(*
SPDX-FileCopyrightText: © 2026 Oleksandr Tiutyk <trofimich@gmail.com>
SPDX-License-Identifier: MIT
License: https://opensource.org/license/mit
*)

(*!
<summary>Checks that a configured task name survives the STOPPED to READY reset.</summary>
<description>
Completes a resource-free one-step task before invoking Reset. A new local fixture is used on every run.
</description>
*)

{attribute 'no_explicit_call' := 'do not call this function block directly'}
FUNCTION_BLOCK TaskNamePreservedByResetTest EXTENDS TOF_Testing.SingleCycleTest
VAR_STAT
	{attribute 'hide'}
	_ClassName : STRING := __POUNAME();
END_VAR

//! <summary>Verifies the constructor name and exercises Reset from STOPPED before checking that name again.</summary>
METHOD PROTECTED ExecuteTest
VAR
	task : CounterTask(name := "Configured counter");
	started : BOOL;
	resetSucceeded : BOOL;
END_VAR
Assert.ThatWideString(actual := task.Name, message := "Task must adopt the explicit constructor name")
	.ToBe(expected := "Configured counter");

task.TargetValue := 1;
started := task.Start();
Assert.ThatBool(actual := started, message := "Fixture must accept Start").IsTrue();

IF NOT started THEN
	RETURN;
END_IF

task.Execute();
Assert.ThatBool(actual := task.State.Stopped, message := "Reset test requires a completed task").IsTrue();

IF NOT task.State.Stopped THEN
	RETURN;
END_IF

resetSucceeded := task.Reset();
Assert.ThatBool(actual := resetSucceeded, message := "Fixture must accept Reset from STOPPED").IsTrue();
Assert.ThatBool(actual := task.State.Ready, message := "Reset must return the fixture to READY").IsTrue();
Assert.ThatWideString(actual := task.Name, message := "Reset from STOPPED must preserve the configured name")
	.ToBe(expected := "Configured counter");
END_METHOD

//! <summary>Borrows the concrete class name. Callers must not modify the returned storage.</summary>
{attribute 'monitoring' := 'call'}
PROPERTY ClassName : REFERENCE TO STRING
GET
ClassName REF= _ClassName;
END_GET
END_PROPERTY

//! <summary>Borrows the compiler-initialized namespace name. Callers must not modify the returned storage.</summary>
{attribute 'monitoring' := 'call'}
PROPERTY NamespaceName : REFERENCE TO STRING
GET
NamespaceName REF= CurrentNamespace.Name;
END_GET
END_PROPERTY

//! <summary>Reports the complete concrete instance size in bytes.</summary>
{attribute 'monitoring' := 'call'}
PROPERTY SelfSize : ULINT
GET
SelfSize := XSIZEOF(THIS^);
END_GET
END_PROPERTY

END_FUNCTION_BLOCK

(* stored: Version 1.1.0.1
   POU TaskNamePreservedByResetTest: Id {5b39e737-dff4-413a-a0dd-cd25526cac07}, SpecialFunc None
   Method ExecuteTest: Id {52b042a6-628e-4f71-a29b-019c5134155c}
   Property ClassName: Id {6afd0256-1dbb-4b5c-9861-094d7b76e291}
   Get Get: Id {31f25c84-b4c1-485a-991b-4dc88ea39adc}
   Property NamespaceName: Id {493fd736-8145-4151-9bfb-b9a7e8e72058}
   Get Get: Id {f789b37c-dce0-468b-88e4-433e87238705}
   Property SelfSize: Id {210b992b-bd78-42eb-9784-5896302ad9fc}
   Get Get: Id {f2cad7d1-93cd-4ac0-9aad-b7d7730204a7} *)
